(* LS Electric XG5000 project: NewProject *)
(* PLC LSPLC *)

PROGRAM NewProgram (* task: 스캔 프로그램 *)
%MX0 := TRUE;
END_PROGRAM